// TIA Portal V21 export
// export: Created 2026-08-21T20:18:53.7310443Z, ExportSetting None, DisplayName Totally Integrated Automation Portal, DisplayVersion V21, DisplayName STEP 7 Professional, DisplayVersion V21, DisplayName STEP 7 Safety, DisplayVersion V21, DisplayName Tech WebApplication, DisplayVersion V21, DisplayName WinCC Basic/Comfort/Advanced, DisplayVersion V21, DisplayName WinCC Professional, DisplayVersion V21, DisplayName WinCC Unified, DisplayVersion V21
FUNCTION_BLOCK "MTPMonBinDrv_Type1"   // FB13, FBD
{ S7_Optimized_Access := 'TRUE' }
// stored: MemoryReserve 100, SetENOAutomatically false
   VAR_INPUT
      from_Ctrl { ExternalAccessible := 'False'; ExternalVisible := 'False'; ExternalWritable := 'False'} : "StruCm";
      Service_Occupied { ExternalAccessible := 'False'; ExternalVisible := 'False'; ExternalWritable := 'False'} : Bool;
      Cmd_Auto { ExternalAccessible := 'False'; ExternalVisible := 'False'; ExternalWritable := 'False'} : Bool;
      Cmd_Man { ExternalAccessible := 'False'; ExternalVisible := 'False'; ExternalWritable := 'False'} : Bool;
      Cmd_StartAut { ExternalAccessible := 'False'; ExternalVisible := 'False'; ExternalWritable := 'False'} : Bool;
      Cmd_StopAut { ExternalAccessible := 'False'; ExternalVisible := 'False'; ExternalWritable := 'False'} : Bool;
      Cmd_Reset { ExternalAccessible := 'False'; ExternalVisible := 'False'; ExternalWritable := 'False'} : Bool;
      PV_In : Bool;
      Intlk04_In01 { ExternalAccessible := 'False'; ExternalVisible := 'False'; ExternalWritable := 'False'} : "DigVal";
      Intlk04_InvIn01 : Bool;
      Intlk04_In1String : String;
      Intlk04_In02 { ExternalAccessible := 'False'; ExternalVisible := 'False'; ExternalWritable := 'False'} : "DigVal";
      Intlk04_InvIn02 : Bool;
      Intlk04_In2String { ExternalAccessible := 'False'; ExternalVisible := 'False'; ExternalWritable := 'False'} : String;
      Intlk04_In03 { ExternalAccessible := 'False'; ExternalVisible := 'False'; ExternalWritable := 'False'} : "DigVal";
      Intlk04_InvIn03 : Bool;
      Intlk04_In3String { ExternalAccessible := 'False'; ExternalVisible := 'False'; ExternalWritable := 'False'} : String;
      Intlk04_In04 { ExternalAccessible := 'False'; ExternalVisible := 'False'; ExternalWritable := 'False'} : "DigVal";
      Intlk04_InvIn04 : Bool;
      Intlk04_In4String { ExternalAccessible := 'False'; ExternalVisible := 'False'; ExternalWritable := 'False'} : String;
   END_VAR
   VAR_OUTPUT
      to_Ctrl { ExternalAccessible := 'False'; ExternalVisible := 'False'; ExternalWritable := 'False'} : "StruCm";
      Occupied { ExternalAccessible := 'False'; ExternalVisible := 'False'; ExternalWritable := 'False'} : Bool;   // Occupied by a Service procedure
      AutAct { ExternalAccessible := 'False'; ExternalVisible := 'False'; ExternalWritable := 'False'} : Bool;
      ManAct { ExternalAccessible := 'False'; ExternalVisible := 'False'; ExternalWritable := 'False'} : Bool;
      PV_Out { ExternalAccessible := 'False'; ExternalVisible := 'False'; ExternalWritable := 'False'} : Bool;
      FbkRunOut : Bool;
      RunOut : Bool;
      Stop { ExternalAccessible := 'False'; ExternalVisible := 'False'; ExternalWritable := 'False'} : Bool;
      GrpErr { ExternalAccessible := 'False'; ExternalVisible := 'False'; ExternalWritable := 'False'} : Bool;
   END_VAR
   VAR
      ChOut { S7_SetPoint := 'True'} : "DiOu";
      DiChIn { S7_SetPoint := 'True'} : "DiIn";
      Intlk04_IDB : "Intlk04";
      MotL_IDB { S7_SetPoint := 'True'} : "MotL";
      MTPMonBinDrv_IDB { ExternalVisible := 'False'; S7_SetPoint := 'True'} : "MTPMonBinDrv";
   END_VAR
   VAR_TEMP
      Intlock : "DigVal";
      CSF_NOP : "DigVal";
      BadOut : "DigVal";
      InverterBad : "DigVal";
      FbkRun : "DigVal";
   END_VAR
   // Intlk04_In01.Value := true;
   // Intlk04_In02.Value := true;
   // Intlk04_In03.Value := true;
   // Intlk04_In04.Value := true;
BEGIN

REGION Network 1: Mod switch
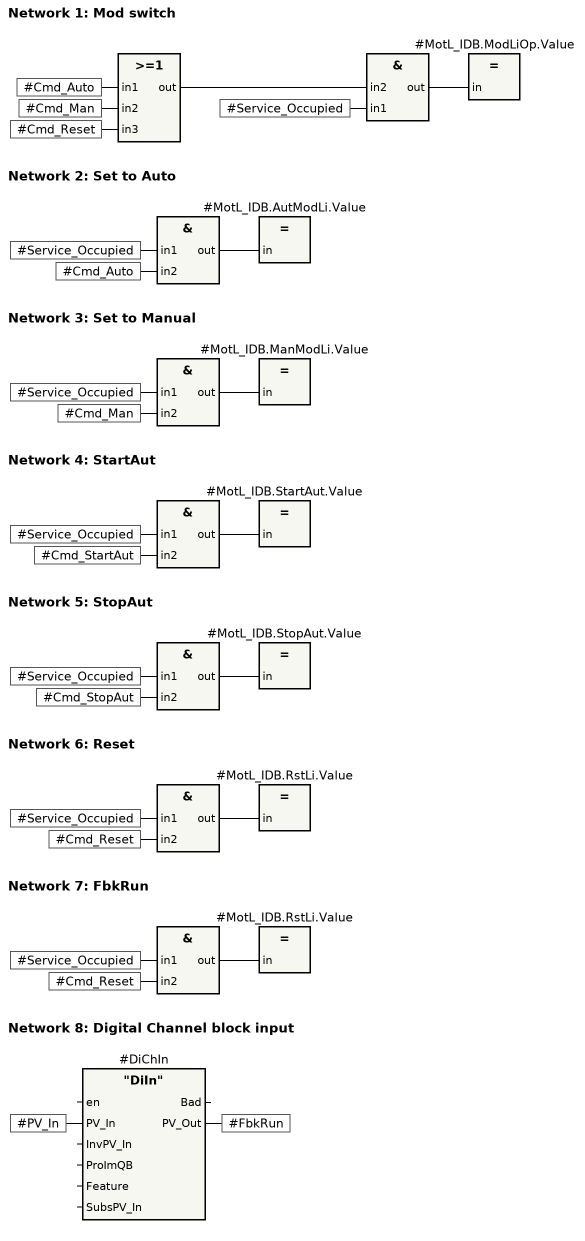
   #MotL_IDB.ModLiOp.Value := (#Cmd_Auto OR #Cmd_Man OR #Cmd_Reset) AND #Service_Occupied;
END_REGION

REGION Network 2: Set to Auto
   #MotL_IDB.AutModLi.Value := #Service_Occupied AND #Cmd_Auto;
END_REGION

REGION Network 3: Set to Manual
   #MotL_IDB.ManModLi.Value := #Service_Occupied AND #Cmd_Man;
END_REGION

REGION Network 4: StartAut
   #MotL_IDB.StartAut.Value := #Service_Occupied AND #Cmd_StartAut;
END_REGION

REGION Network 5: StopAut
   #MotL_IDB.StopAut.Value := #Service_Occupied AND #Cmd_StopAut;
END_REGION

REGION Network 6: Reset
   #MotL_IDB.RstLi.Value := #Service_Occupied AND #Cmd_Reset;
END_REGION

REGION Network 7: FbkRun
   #MotL_IDB.RstLi.Value := #Service_Occupied AND #Cmd_Reset;
END_REGION

REGION Network 8: Digital Channel block input
   #DiChIn(PV_In := #PV_In, PV_Out => #FbkRun);   // "DiIn"
END_REGION

REGION Network 9: CSF
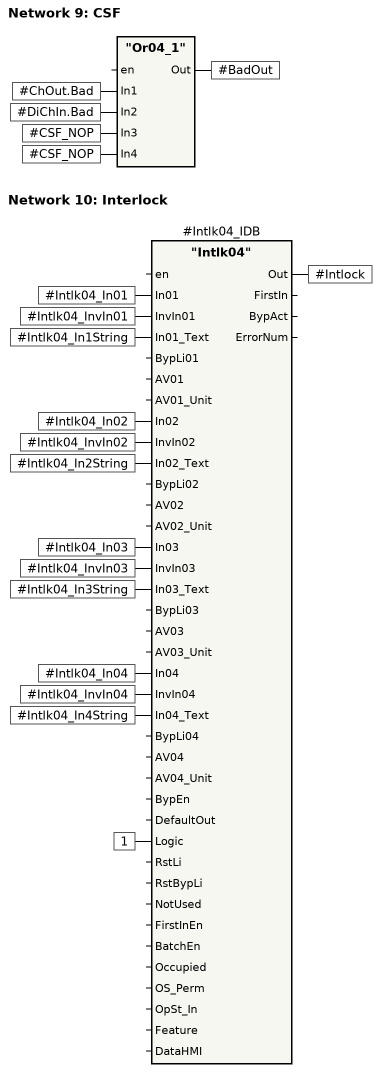
   "Or04_1"(In1 := #ChOut.Bad, In2 := #DiChIn.Bad, In3 := #CSF_NOP, In4 := #CSF_NOP, Out => #BadOut);
END_REGION

REGION Network 10: Interlock
   #Intlk04_IDB(In01 := #Intlk04_In01,   // "Intlk04"
                InvIn01 := #Intlk04_InvIn01,
                In01_Text := #Intlk04_In1String,
                In02 := #Intlk04_In02,
                InvIn02 := #Intlk04_InvIn02,
                In02_Text := #Intlk04_In2String,
                In03 := #Intlk04_In03,
                InvIn03 := #Intlk04_InvIn03,
                In03_Text := #Intlk04_In3String,
                In04 := #Intlk04_In04,
                InvIn04 := #Intlk04_InvIn04,
                In04_Text := #Intlk04_In4String,
                Logic := 1,
                Out => #Intlock);
END_REGION

REGION Network 11: MotSpdCL
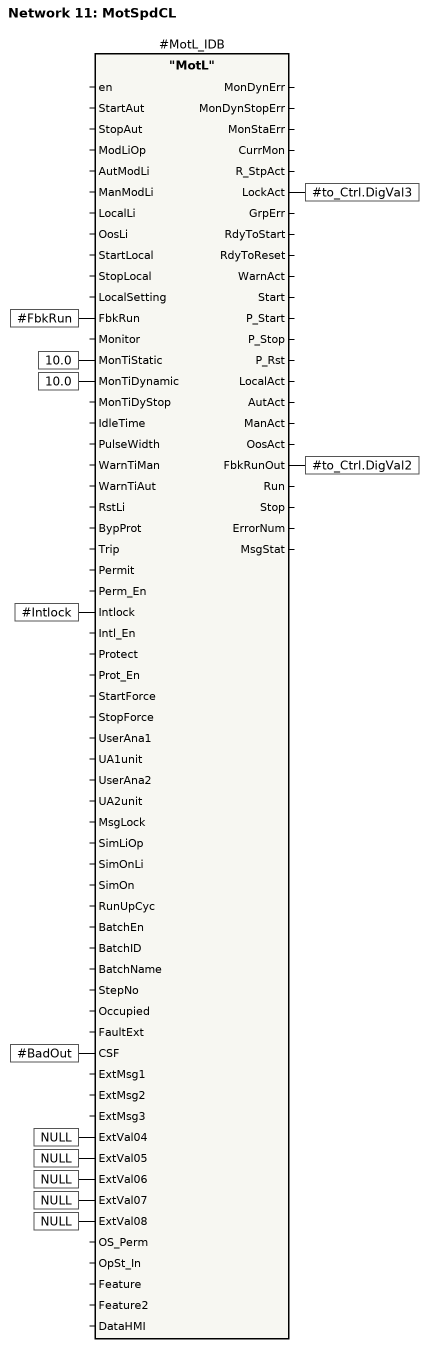
   #MotL_IDB(FbkRun := #FbkRun,   // "MotL"
             MonTiStatic := 10.0,
             MonTiDynamic := 10.0,
             Intlock := #Intlock,
             CSF := #BadOut,
             ExtVal04 := NULL,
             ExtVal05 := NULL,
             ExtVal06 := NULL,
             ExtVal07 := NULL,
             ExtVal08 := NULL,
             LockAct => #to_Ctrl.DigVal3,
             FbkRunOut => #to_Ctrl.DigVal2);
END_REGION

REGION Network 12: Channel block output
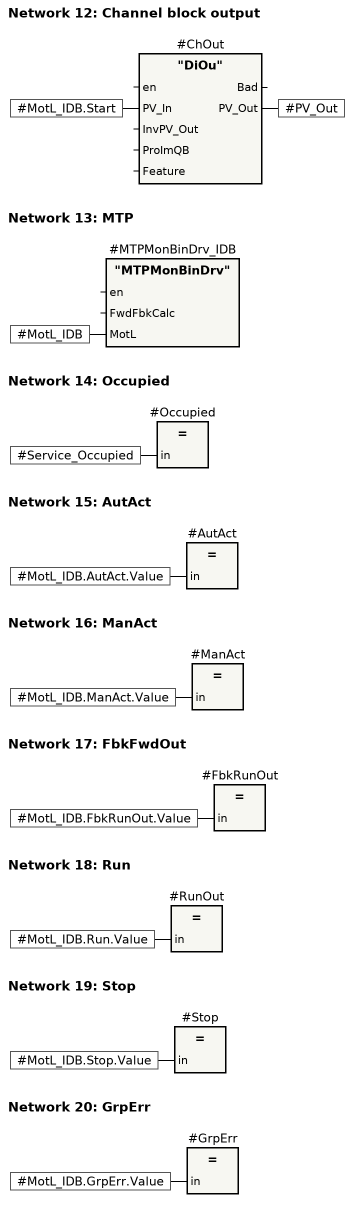
   #ChOut(PV_In := #MotL_IDB.Start, PV_Out => #PV_Out);   // "DiOu"
END_REGION

REGION Network 13: MTP
   #MTPMonBinDrv_IDB(MotL := #MotL_IDB);   // "MTPMonBinDrv"
END_REGION

REGION Network 14: Occupied
   #Occupied := #Service_Occupied;
END_REGION

REGION Network 15: AutAct
   #AutAct := #MotL_IDB.AutAct.Value;
END_REGION

REGION Network 16: ManAct
   #ManAct := #MotL_IDB.ManAct.Value;
END_REGION

REGION Network 17: FbkFwdOut
   #FbkRunOut := #MotL_IDB.FbkRunOut.Value;
END_REGION

REGION Network 18: Run
   #RunOut := #MotL_IDB.Run.Value;
END_REGION

REGION Network 19: Stop
   #Stop := #MotL_IDB.Stop.Value;
END_REGION

REGION Network 20: GrpErr
   #GrpErr := #MotL_IDB.GrpErr.Value;
END_REGION
END_FUNCTION_BLOCK
